(* IEC 61131-3 sources: codesys-framework/txt/application/ToDo/Utils/FB_GetIpAddress, 2 files *)

(* ---- GetAddress.method.st ---- *)
METHOD GetAddress : STRING
VAR_INPUT
END_VAR

// --- BEGIN IMPLEMENTATION ---

GetAddress := _sIp;

(* ---- ReadAddress.method.st ---- *)
METHOD ReadAddress
VAR_INPUT
END_VAR

// --- BEGIN IMPLEMENTATION ---

_xRead := TRUE;
